PROGRAM Gr00Home
VAR_INPUT
	(* Input variables / Eingang Variablen *)
	bEnable					:BOOL;						(* Enable Gr00Home *)
	bExecute				:BOOL;						(* Home execute *)

	(* Instances *)
	fbInit						:FB_Gr00HomeInit;
	fbProcedure				:FB_Gr00HomeProcedure;
END_VAR
VAR
	(* Enummerations *)

	(* Variables *)

	(* References *)

	(* Interfaces *)

	(* Instances *)
	rtExecute					:R_TRIG;

	fbAlarm					:FB_Gr00HomeAlarm;

END_VAR
VAR CONSTANT
	nFatalErrorMaxIdx				:INT := 0;						(* Maximal index of  using alarms *)
	nErrorMaxIdx					:INT := 0;						(* Maximal index of  using alarms *)
	nWarningMaxIdx				:INT := 0;						(* Maximal index of  using alarms *)
	nMessageMaxIdx				:INT := 0;						(* Maximal index of  using alarms *)
	nHintMaxIdx					:INT := 0;						(* Maximal index of  using alarms *)

	dnFatalErrorBaseIdentNo		:DINT := 03000;				(* Fatal error identification number *)
	dnErrorBaseIdentNo			:DINT := 03100;				(* Error identification number *)
	dnWarningBaseIdentNo		:DINT := 03200;				(* Warning identification number *)
	dnMessageBaseIdentNo		:DINT := 03300;				(* Message identification number *)
	dnHintBaseIdentNo			:DINT := 03400;				(* Hint identification number *)
END_VAR

IF NOT bEnable
THEN
	RETURN;
END_IF;

(* Check home execute *)
bExecute := etgGr00MachineState = ET_MachineState_eHomeRefExe
		      OR etgGr00MachineState = ET_MachineState_eHomeExe;

rtExecute(CLK := bExecute);                   

IF rtExecute.Q
THEN
	fbInit.bFirstTime := FALSE;
	A_Init();
END_IF;

A_Procedure();
A_Alarm();

ACTION A_Alarm:

(* Collect and execute input alarms *)
fbAlarm.stAlarmIn.arbError[0].bActive := fbProcedure.bErrorByProgramVerification;
fbAlarm.stAlarmIn.arbError[0].dnCode := dnErrorBaseIdentNo + 0;

fbAlarm(
	etMachineMode := etgGr00MachineMode,
	etMachineState := etgGr00MachineState,
	bNoEStop := bgGr00NoEmergencyStop,
	bConfirmAlarm := bgGr00ConfirmAlarm,
	dtDateTime := stgGr00DateTime.dtDateTime,
	nFatalErrorMaxIdx := nFatalErrorMaxIdx,
	nErrorMaxIdx := nErrorMaxIdx,
	nWarningMaxIdx := nWarningMaxIdx,
	nMessageMaxIdx := nMessageMaxIdx,
	nHintMaxIdx := nHintMaxIdx,
	bMoveInterrupted := bgGr00MoveInterrupted,
	bHomeCompleted := bgGr00HomeCompleted,
	stAlarmOut => stgGr00Alarm.stHome
);
END_ACTION

ACTION A_Init:

(* Initializing variables *)
fbInit();
END_ACTION

ACTION A_Procedure:

(* Execute home procedure *)
fbProcedure(
	bEnable := etgGr00MachineMode = ET_MachineMode_eHome,
	bExecute := rtExecute.Q,
	bReleaseNextStep := etgGr00MachineState = ET_MachineState_eHomeRefExe
		      	     		      OR etgGr00MachineState = ET_MachineState_eHomeExe
);
END_ACTION

END_PROGRAM

(* stored: Version 1.1.0.1, ProductVersion 3.1.4024.15
   POU Gr00Home: Id {5c2522d3-964b-4903-b6ed-f457f697d2f7}, SpecialFunc None
   Action A_Alarm: Id {1ea6b778-9874-4754-87db-6526503c9c77}
   Action A_Init: Id {b7245eca-8ce4-4698-860c-d232020376a9}
   Action A_Procedure: Id {9fec207b-2d67-4d32-9dcf-0fcf2642d203} *)
